(* PLC project Vn_targets_after_box, Beckhoff Automation GmbH TwinCAT PLC Control 3.5.13.21 *)
(* stored: creationDateTime 1970-01-01T00:00:00 *)

PROGRAM Vn_targets_after_box
  VAR  (* added by the conversion: wires and edge detectors of the diagram *)
    _OR10000000007_OUT : BOOL;
  END_VAR

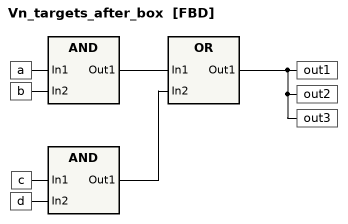
(* FBD diagram, written out as Structured Text *)
_OR10000000007_OUT := a AND b OR c AND d;
out1 := _OR10000000007_OUT;
out2 := _OR10000000007_OUT;
out3 := _OR10000000007_OUT;
END_PROGRAM
